Omron CX-Programmer project NewProject (CX-Programmer 9.61)

# PLC NewPLC1: CJ1H-H CPU65
I/O table (CPU CJ1M-CPU21): rack 0 slot 0 CJ1W-ETN21(ETN21Mode); rack 0 slot 1 CJ1W-DRM21; rack 0 slot 2 CJ1W-ID211; rack 0 slot 3 CJ1W-ID211; rack 0 slot 4 CJ1W-ID211; rack 0 slot 5 CJ1W-OD211; rack 0 slot 6 CJ1W-OD212; rack 0 slot 7 CJ1W-OC211; rack 0 slot 8 CJ1W-MAD42

## Global symbols (name address type ; comment)
W4.01 BOOL  ; Лифт №1 РЕЛЕ ВКЛ питание
W5.01 BOOL  ; Лифт №1 Реле выкл Питание
BLINK_L1 BLINK
BLINK_L2 BLINK  ; Сигнализация не готовности лифта
DOWN W1.03 BOOL
DOWN_stop W0.03 BOOL
HOME_L1 W0.08 BOOL  ; Лифт откальброван
L1_DOWN W0.00 BOOL
L1_UP W0.01 BOOL
L2_DOWN W0.04 BOOL
L2_DOWN_stop W0.07 BOOL
L2_UP W0.05 BOOL
L2_UP_stop W0.06 BOOL
ON W1.00 BOOL
UP W1.02 BOOL
UP_stop W0.02 BOOL

## Program MotorDrive_LIFT_1 (cyclic task 0)
Local symbols
BLINK_1_OUT W1.01 BOOL
L1_Key_start 0.08 BOOL  ; $?St$Bk?_#[231] / Лифт №1 Кнопка "Старт"$?St$Bk?_#[231]
L1_Key_stop 0.09 BOOL  ; $?St$Bk?_#[232] / Лифт №1 Кнопка "Стоп"$?St$Bk?_#[232]
L1_Lamp_start 3.06 BOOL  ; Лифт №1 Лампа Старт
L1_in_N_limit 1.06 BOOL  ; Лифт №1 Нижний аварийный концевик
L1_in_P_limit 1.07 BOOL  ; Лифт №1 Верхний аварийный концевик
L1_out_Down 4.08 BOOL  ; Лифт №1 Реле ВКЛ движение вниз
L1_out_Drag 4.12 BOOL  ; Лифт №1 Реле отключение тормоза
L1_out_Up 4.10 BOOL  ; Лифт №1 Реле ВКЛ движение вверх
L1_out_powerON 4.14 BOOL  ; Лифт №1 Реле ВКЛ питание

### Section POWER

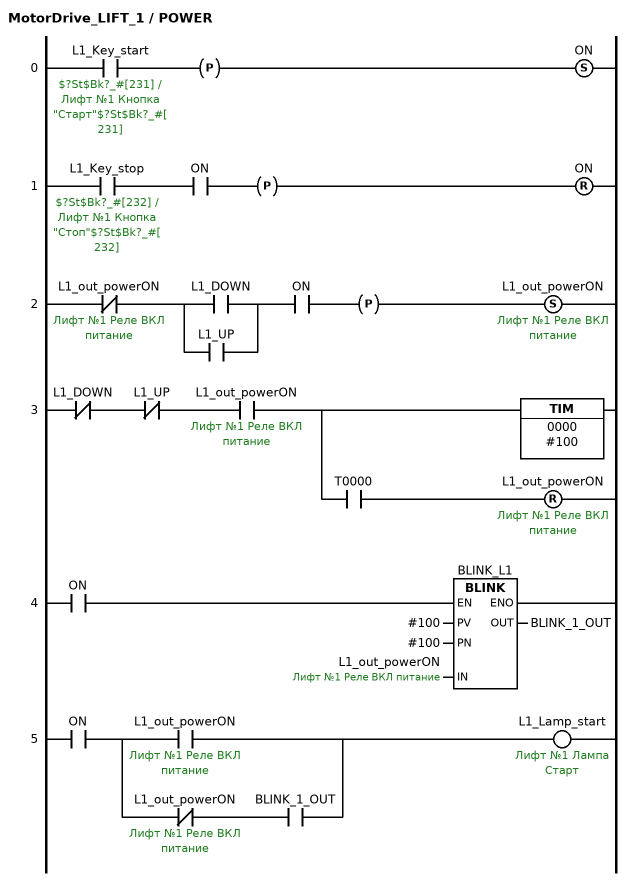
; rung 0
LD L1_Key_start  ; $?St$Bk?_#[231] / Лифт №1 Кнопка "Старт"$?St$Bk?_#[231]
UP(521)
SET ON
; rung 1
LD L1_Key_stop  ; $?St$Bk?_#[232] / Лифт №1 Кнопка "Стоп"$?St$Bk?_#[232]
AND ON
UP(521)
RSET ON
; rung 2
LDNOT L1_out_powerON  ; Лифт №1 Реле ВКЛ питание
LD L1_DOWN
OR L1_UP
ANDLD
AND ON
UP(521)
SET L1_out_powerON  ; Лифт №1 Реле ВКЛ питание
; rung 3
LDNOT L1_DOWN
ANDNOT L1_UP
AND L1_out_powerON  ; Лифт №1 Реле ВКЛ питание
TIM 0000 #100
AND T0000
RSET L1_out_powerON  ; Лифт №1 Реле ВКЛ питание
; rung 4
LD ON
CALL BLINK_L1 : BLINK (PV := #100, PN := #100, IN := L1_out_powerON, OUT => BLINK_1_OUT)  ; Лифт №1 Реле ВКЛ питание
; rung 5
LD ON
LD L1_out_powerON  ; Лифт №1 Реле ВКЛ питание
LDNOT L1_out_powerON  ; Лифт №1 Реле ВКЛ питание
AND BLINK_1_OUT
ORLD
ANDLD
OUT L1_Lamp_start  ; Лифт №1 Лампа Старт

### Section UP

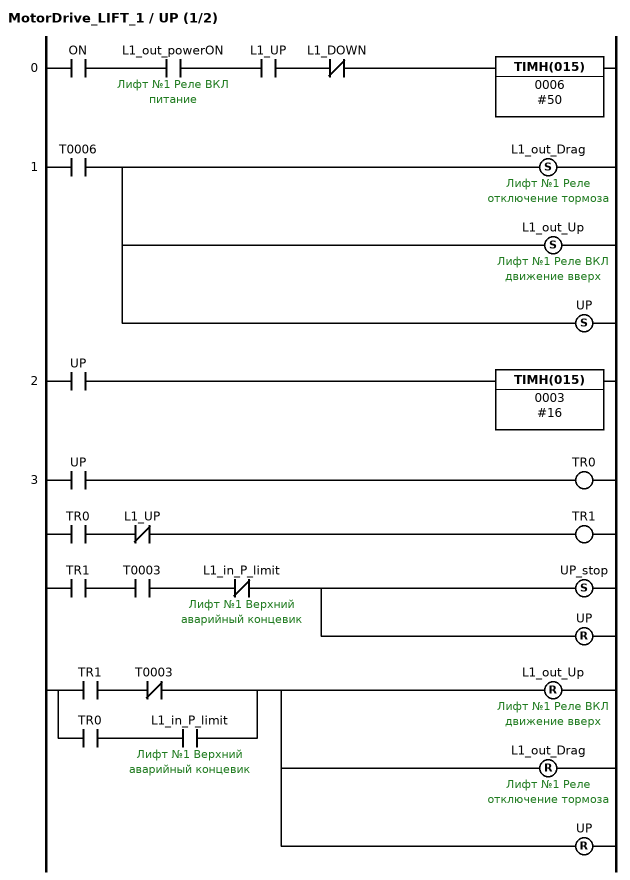
; rung 0
LD ON
AND L1_out_powerON  ; Лифт №1 Реле ВКЛ питание
AND L1_UP
ANDNOT L1_DOWN
TIMH(015) 0006 #50
; rung 1
LD T0006
SET L1_out_Drag  ; Лифт №1 Реле отключение тормоза
SET L1_out_Up  ; Лифт №1 Реле ВКЛ движение вверх
SET UP
; rung 2
LD UP
TIMH(015) 0003 #16
; rung 3
LD UP
OUT TR0
ANDNOT L1_UP
OUT TR1
AND T0003
ANDNOT L1_in_P_limit  ; Лифт №1 Верхний аварийный концевик
SET UP_stop
RSET UP
LD TR1
ANDNOT T0003
LD TR0
AND L1_in_P_limit  ; Лифт №1 Верхний аварийный концевик
ORLD
RSET L1_out_Up  ; Лифт №1 Реле ВКЛ движение вверх
RSET L1_out_Drag  ; Лифт №1 Реле отключение тормоза
RSET UP

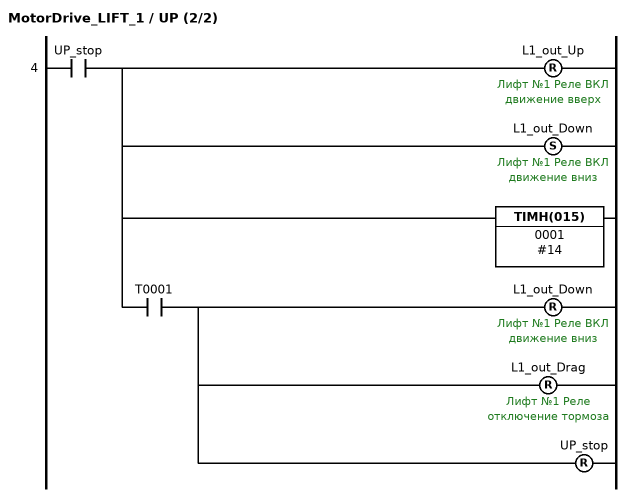
; rung 4
LD UP_stop
RSET L1_out_Up  ; Лифт №1 Реле ВКЛ движение вверх
SET L1_out_Down  ; Лифт №1 Реле ВКЛ движение вниз
TIMH(015) 0001 #14
AND T0001
RSET L1_out_Down  ; Лифт №1 Реле ВКЛ движение вниз
RSET L1_out_Drag  ; Лифт №1 Реле отключение тормоза
RSET UP_stop

### Section DOWN

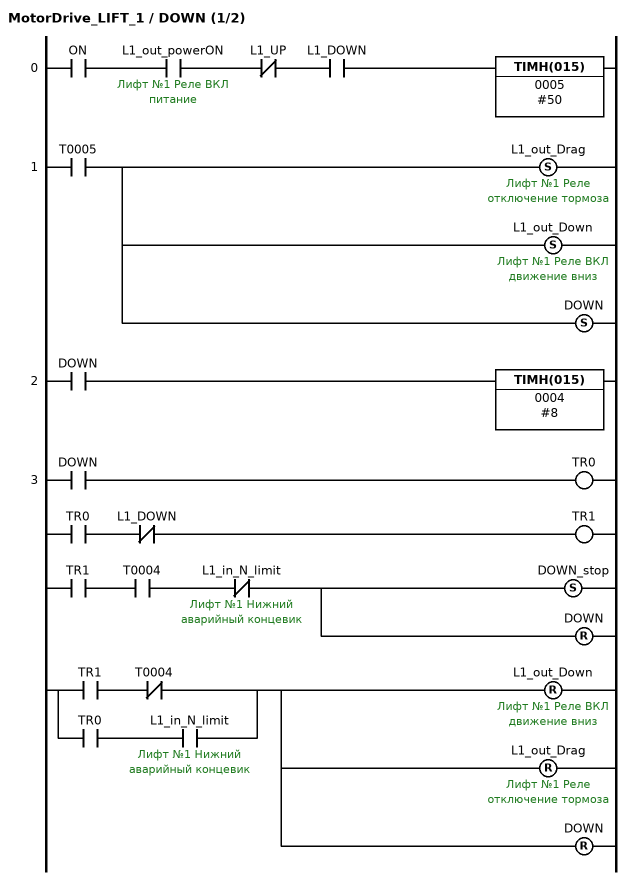
; rung 0
LD ON
AND L1_out_powerON  ; Лифт №1 Реле ВКЛ питание
ANDNOT L1_UP
AND L1_DOWN
TIMH(015) 0005 #50
; rung 1
LD T0005
SET L1_out_Drag  ; Лифт №1 Реле отключение тормоза
SET L1_out_Down  ; Лифт №1 Реле ВКЛ движение вниз
SET DOWN
; rung 2
LD DOWN
TIMH(015) 0004 #8
; rung 3
LD DOWN
OUT TR0
ANDNOT L1_DOWN
OUT TR1
AND T0004
ANDNOT L1_in_N_limit  ; Лифт №1 Нижний аварийный концевик
SET DOWN_stop
RSET DOWN
LD TR1
ANDNOT T0004
LD TR0
AND L1_in_N_limit  ; Лифт №1 Нижний аварийный концевик
ORLD
RSET L1_out_Down  ; Лифт №1 Реле ВКЛ движение вниз
RSET L1_out_Drag  ; Лифт №1 Реле отключение тормоза
RSET DOWN

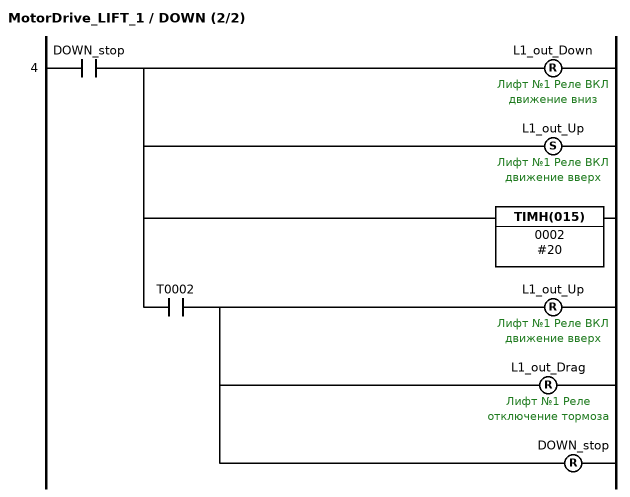
; rung 4
LD DOWN_stop
RSET L1_out_Down  ; Лифт №1 Реле ВКЛ движение вниз
SET L1_out_Up  ; Лифт №1 Реле ВКЛ движение вверх
TIMH(015) 0002 #20
AND T0002
RSET L1_out_Up  ; Лифт №1 Реле ВКЛ движение вверх
RSET L1_out_Drag  ; Лифт №1 Реле отключение тормоза
RSET DOWN_stop

### Section END
; rung 0
END(001)

## Program NewProgram1 (cyclic task 1)
Local symbols
BLINK_2_OUT W2.01 BOOL
F_Key_lev1 2.01 BOOL  ; Этаж 1 Кнопка вызова лифта
F_Key_lev2 2.03 BOOL  ; Этаж 2 Кнопка вызова лифта
F_Key_lev3 2.05 BOOL  ; Этаж 3 Кнопка вызова лифта
F_Key_lev4 2.07 BOOL  ; Этаж 4 Кнопка вызова лифта
F_Key_lev5 2.09 BOOL  ; Этаж 5 Кнопка вызова лифта
F_Key_lev6 2.11 BOOL  ; Этаж 6 Кнопка вызова лифта
HOME_L1_NOT W2.02 BOOL
L1_Key_lev1 0.10 BOOL  ; $?St$Bk?_#[251] / Лифт №1 Кнопка "Этаж 1"$?St$Bk?_#[251]
L1_Key_lev2 0.12 BOOL  ; $?St$Bk?_#[252] / Лифт №1 Кнопка "Этаж 2"$?St$Bk?_#[252]
L1_Key_lev3 0.14 BOOL  ; $?St$Bk?_#[253] / Лифт №1 Кнопка "Этаж 3"$?St$Bk?_#[253]
L1_Key_lev4 0.11 BOOL  ; $?St$Bk?_#[254] / Лифт №1 Кнопка "Этаж 4"$?St$Bk?_#[254]
L1_Key_lev5 0.13 BOOL  ; $?St$Bk?_#[255] / Лифт №1 Кнопка "Этаж 5"$?St$Bk?_#[255]
L1_Key_lev6 0.15 BOOL  ; $?St$Bk?_#[256] / Лифт №1 Кнопка "Этаж 6"$?St$Bk?_#[256]
L1_Lamp_lev1 3.04 BOOL  ; Лифт №1 Лампа Этаж 1
L1_Lamp_lev2 3.02 BOOL  ; Лифт №1 Лампа Этаж 2
L1_Lamp_lev3 3.00 BOOL  ; Лифт №1 Лампа Этаж 3
L1_Lamp_lev4 3.05 BOOL  ; Лифт №1 Лампа Этаж 4
L1_Lamp_lev5 3.03 BOOL  ; Лифт №1 Лампа Этаж 5
L1_Lamp_lev6 3.01 BOOL  ; Лифт №1 Лампа Этаж 6
L1_Lamp_start 3.06 BOOL  ; Лифт №1 Лампа Старт
L1_Lamp_stop 3.07 BOOL  ; Лифт №1 Лампа Стоп
L1_in_Floor_1 1.05 BOOL  ; Лифт №1 Датчик Этаж 1
L1_in_Floor_2 1.04 BOOL  ; Лифт №1 Датчик Этаж 2
L1_in_Floor_3 1.03 BOOL  ; Лифт №1 Датчик Этаж 3
L1_in_Floor_4 1.02 BOOL  ; Лифт №1 Датчик Этаж 4
L1_in_Floor_5 1.01 BOOL  ; Лифт №1 Датчик Этаж 5
L1_in_Floor_6 1.00 BOOL  ; Лифт №1 Датчик Этаж 6
L1_in_N_limit 1.06 BOOL  ; Лифт №1 Нижний аварийный концевик
L1_in_P_limit 1.07 BOOL  ; Лифт №1 Верхний аварийный концевик
L1_out_powerON 4.14 BOOL  ; Лифт №1 Реле ВКЛ питание

### Section HM

### Section Doors

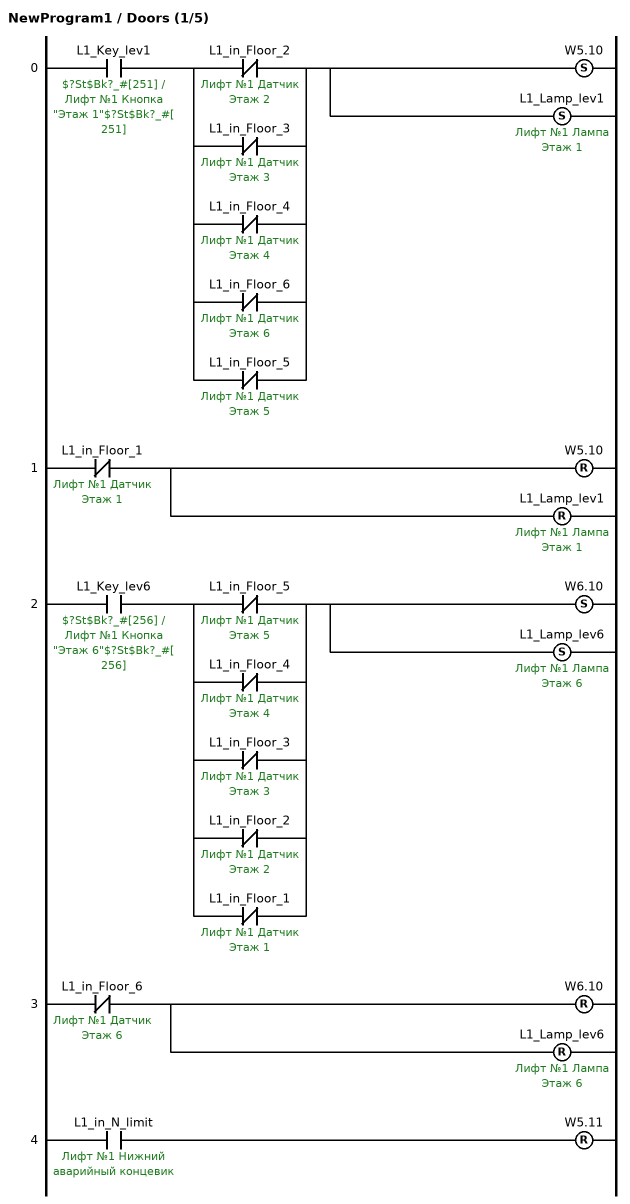
; rung 0
LD L1_Key_lev1  ; $?St$Bk?_#[251] / Лифт №1 Кнопка "Этаж 1"$?St$Bk?_#[251]
LDNOT L1_in_Floor_2  ; Лифт №1 Датчик Этаж 2
ORNOT L1_in_Floor_3  ; Лифт №1 Датчик Этаж 3
ORNOT L1_in_Floor_4  ; Лифт №1 Датчик Этаж 4
ORNOT L1_in_Floor_6  ; Лифт №1 Датчик Этаж 6
ORNOT L1_in_Floor_5  ; Лифт №1 Датчик Этаж 5
ANDLD
SET W5.10
SET L1_Lamp_lev1  ; Лифт №1 Лампа Этаж 1
; rung 1
LDNOT L1_in_Floor_1  ; Лифт №1 Датчик Этаж 1
RSET W5.10
RSET L1_Lamp_lev1  ; Лифт №1 Лампа Этаж 1
; rung 2
LD L1_Key_lev6  ; $?St$Bk?_#[256] / Лифт №1 Кнопка "Этаж 6"$?St$Bk?_#[256]
LDNOT L1_in_Floor_5  ; Лифт №1 Датчик Этаж 5
ORNOT L1_in_Floor_4  ; Лифт №1 Датчик Этаж 4
ORNOT L1_in_Floor_3  ; Лифт №1 Датчик Этаж 3
ORNOT L1_in_Floor_2  ; Лифт №1 Датчик Этаж 2
ORNOT L1_in_Floor_1  ; Лифт №1 Датчик Этаж 1
ANDLD
SET W6.10
SET L1_Lamp_lev6  ; Лифт №1 Лампа Этаж 6
; rung 3
LDNOT L1_in_Floor_6  ; Лифт №1 Датчик Этаж 6
RSET W6.10
RSET L1_Lamp_lev6  ; Лифт №1 Лампа Этаж 6
; rung 4
LD L1_in_N_limit  ; Лифт №1 Нижний аварийный концевик
RSET W5.11

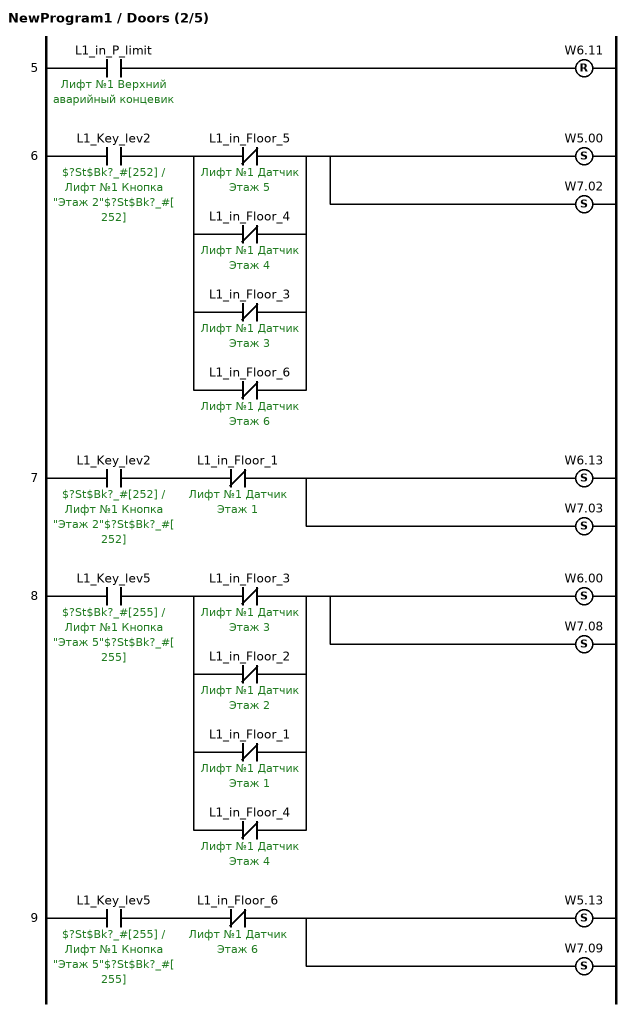
; rung 5
LD L1_in_P_limit  ; Лифт №1 Верхний аварийный концевик
RSET W6.11
; rung 6
LD L1_Key_lev2  ; $?St$Bk?_#[252] / Лифт №1 Кнопка "Этаж 2"$?St$Bk?_#[252]
LDNOT L1_in_Floor_5  ; Лифт №1 Датчик Этаж 5
ORNOT L1_in_Floor_4  ; Лифт №1 Датчик Этаж 4
ORNOT L1_in_Floor_3  ; Лифт №1 Датчик Этаж 3
ORNOT L1_in_Floor_6  ; Лифт №1 Датчик Этаж 6
ANDLD
SET W5.00
SET W7.02
; rung 7
LD L1_Key_lev2  ; $?St$Bk?_#[252] / Лифт №1 Кнопка "Этаж 2"$?St$Bk?_#[252]
ANDNOT L1_in_Floor_1  ; Лифт №1 Датчик Этаж 1
SET W6.13
SET W7.03
; rung 8
LD L1_Key_lev5  ; $?St$Bk?_#[255] / Лифт №1 Кнопка "Этаж 5"$?St$Bk?_#[255]
LDNOT L1_in_Floor_3  ; Лифт №1 Датчик Этаж 3
ORNOT L1_in_Floor_2  ; Лифт №1 Датчик Этаж 2
ORNOT L1_in_Floor_1  ; Лифт №1 Датчик Этаж 1
ORNOT L1_in_Floor_4  ; Лифт №1 Датчик Этаж 4
ANDLD
SET W6.00
SET W7.08
; rung 9
LD L1_Key_lev5  ; $?St$Bk?_#[255] / Лифт №1 Кнопка "Этаж 5"$?St$Bk?_#[255]
ANDNOT L1_in_Floor_6  ; Лифт №1 Датчик Этаж 6
SET W5.13
SET W7.09

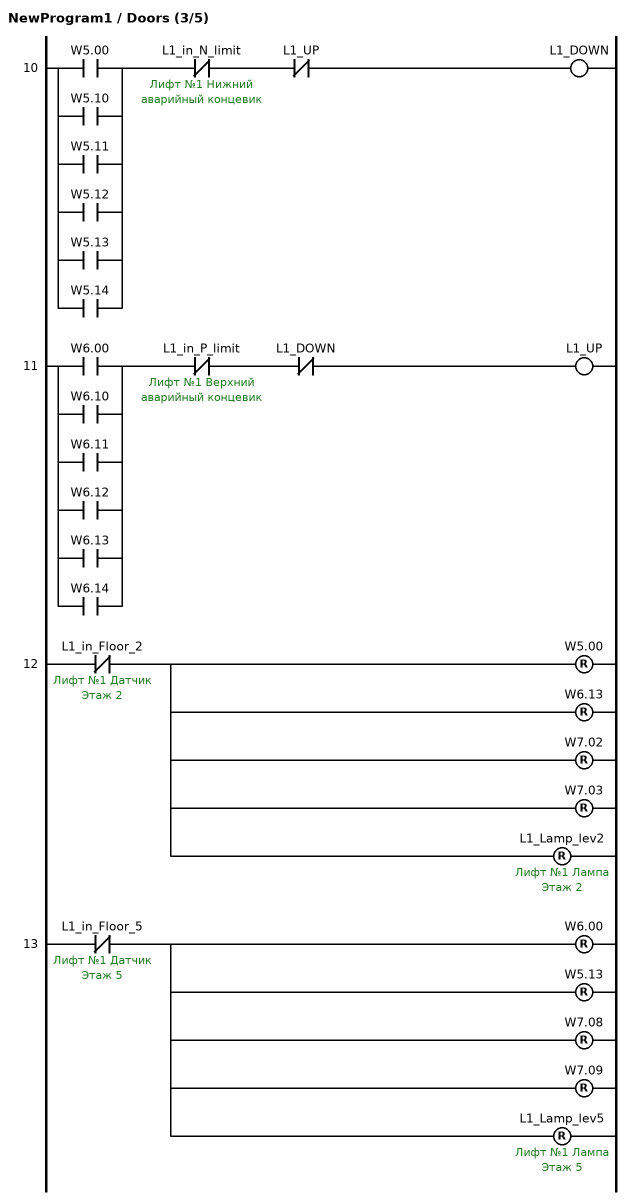
; rung 10
LD W5.00
OR W5.10
OR W5.11
OR W5.12
OR W5.13
OR W5.14
ANDNOT L1_in_N_limit  ; Лифт №1 Нижний аварийный концевик
ANDNOT L1_UP
OUT L1_DOWN
; rung 11
LD W6.00
OR W6.10
OR W6.11
OR W6.12
OR W6.13
OR W6.14
ANDNOT L1_in_P_limit  ; Лифт №1 Верхний аварийный концевик
ANDNOT L1_DOWN
OUT L1_UP
; rung 12
LDNOT L1_in_Floor_2  ; Лифт №1 Датчик Этаж 2
RSET W5.00
RSET W6.13
RSET W7.02
RSET W7.03
RSET L1_Lamp_lev2  ; Лифт №1 Лампа Этаж 2
; rung 13
LDNOT L1_in_Floor_5  ; Лифт №1 Датчик Этаж 5
RSET W6.00
RSET W5.13
RSET W7.08
RSET W7.09
RSET L1_Lamp_lev5  ; Лифт №1 Лампа Этаж 5

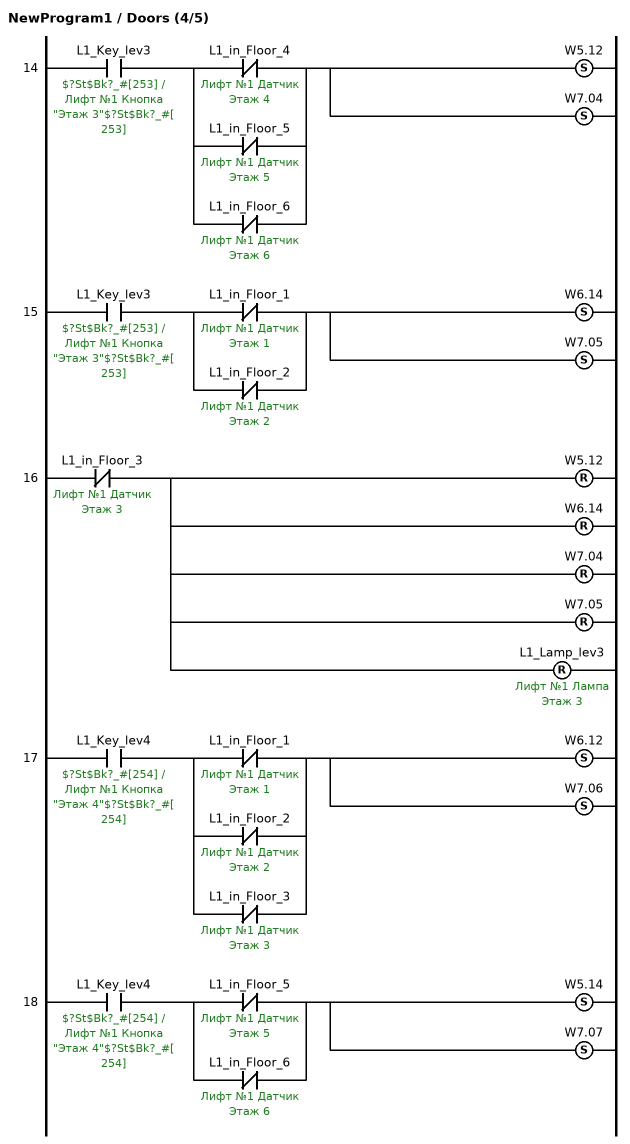
; rung 14
LD L1_Key_lev3  ; $?St$Bk?_#[253] / Лифт №1 Кнопка "Этаж 3"$?St$Bk?_#[253]
LDNOT L1_in_Floor_4  ; Лифт №1 Датчик Этаж 4
ORNOT L1_in_Floor_5  ; Лифт №1 Датчик Этаж 5
ORNOT L1_in_Floor_6  ; Лифт №1 Датчик Этаж 6
ANDLD
SET W5.12
SET W7.04
; rung 15
LD L1_Key_lev3  ; $?St$Bk?_#[253] / Лифт №1 Кнопка "Этаж 3"$?St$Bk?_#[253]
LDNOT L1_in_Floor_1  ; Лифт №1 Датчик Этаж 1
ORNOT L1_in_Floor_2  ; Лифт №1 Датчик Этаж 2
ANDLD
SET W6.14
SET W7.05
; rung 16
LDNOT L1_in_Floor_3  ; Лифт №1 Датчик Этаж 3
RSET W5.12
RSET W6.14
RSET W7.04
RSET W7.05
RSET L1_Lamp_lev3  ; Лифт №1 Лампа Этаж 3
; rung 17
LD L1_Key_lev4  ; $?St$Bk?_#[254] / Лифт №1 Кнопка "Этаж 4"$?St$Bk?_#[254]
LDNOT L1_in_Floor_1  ; Лифт №1 Датчик Этаж 1
ORNOT L1_in_Floor_2  ; Лифт №1 Датчик Этаж 2
ORNOT L1_in_Floor_3  ; Лифт №1 Датчик Этаж 3
ANDLD
SET W6.12
SET W7.06
; rung 18
LD L1_Key_lev4  ; $?St$Bk?_#[254] / Лифт №1 Кнопка "Этаж 4"$?St$Bk?_#[254]
LDNOT L1_in_Floor_5  ; Лифт №1 Датчик Этаж 5
ORNOT L1_in_Floor_6  ; Лифт №1 Датчик Этаж 6
ANDLD
SET W5.14
SET W7.07

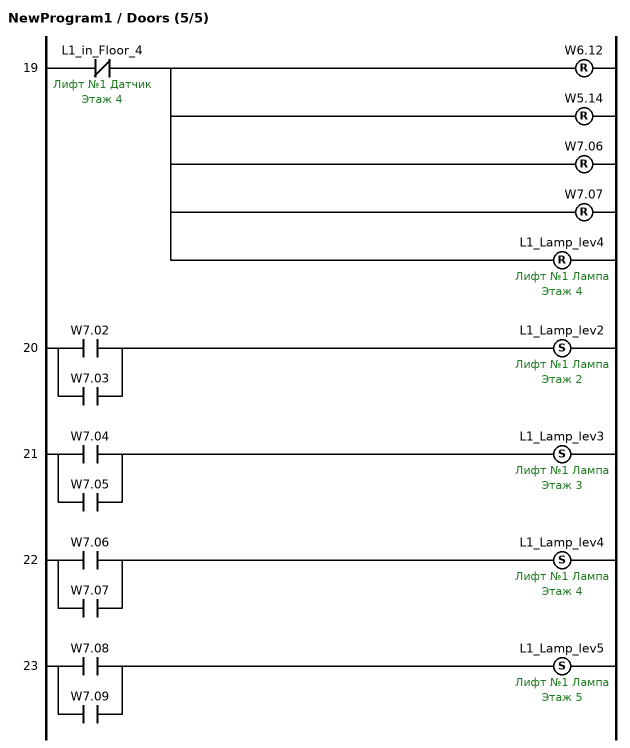
; rung 19
LDNOT L1_in_Floor_4  ; Лифт №1 Датчик Этаж 4
RSET W6.12
RSET W5.14
RSET W7.06
RSET W7.07
RSET L1_Lamp_lev4  ; Лифт №1 Лампа Этаж 4
; rung 20
LD W7.02
OR W7.03
SET L1_Lamp_lev2  ; Лифт №1 Лампа Этаж 2
; rung 21
LD W7.04
OR W7.05
SET L1_Lamp_lev3  ; Лифт №1 Лампа Этаж 3
; rung 22
LD W7.06
OR W7.07
SET L1_Lamp_lev4  ; Лифт №1 Лампа Этаж 4
; rung 23
LD W7.08
OR W7.09
SET L1_Lamp_lev5  ; Лифт №1 Лампа Этаж 5

### Section END
; rung 0
END(001)

## Function block BLINK
VAR_INPUT
  PV : INT;
  PN : INT;
  IN : BOOL;
END_VAR
VAR_OUTPUT
  OUT : BOOL;
END_VAR
VAR
  TIMER_1 : TIMER;
  TIMER_2 : TIMER;
  ON : BOOL;
END_VAR

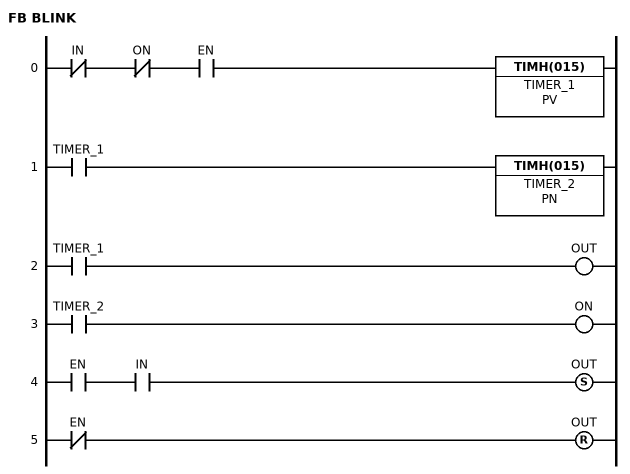
; rung 0
LDNOT IN
ANDNOT ON
AND EN
TIMH(015) TIMER_1 PV
; rung 1
LD TIMER_1
TIMH(015) TIMER_2 PN
; rung 2
LD TIMER_1
OUT OUT
; rung 3
LD TIMER_2
OUT ON
; rung 4
LD EN
AND IN
SET OUT
; rung 5
LDNOT EN
RSET OUT